// TIA Portal V20 export
Screen "Pop-up_Sealer_1"  395x650
  ScreenItem "Robot Name" at 2,2 size 393x48  Type=HmiIOField
  ScreenItem "Background" at -1,49 size 395x601  Type=HmiRectangle
  ScreenItem "Cancel Mode" at 315,4 size 76x42  Type=HmiButton
  ScreenItem "矩形_4" at 31,68 size 324x517  Type=HmiRectangle
  ScreenItem "Text Filed E- Stop_17" at 39,333 size 148x21  Type=HmiTextBox
  ScreenItem "Text Field In Auto On_9" at 39,98 size 148x21  Type=HmiTextBox
  ScreenItem "Text Field Home Position_17" at 39,121 size 148x21  Type=HmiTextBox
  ScreenItem "Text field Robot Status_5" at 33,69 size 324x26  Type=HmiTextBox
  ScreenItem "Text Field Manual_17" at 39,263 size 148x21  Type=HmiTextBox
  ScreenItem "Text Field System Ready_9" at 39,145 size 148x21  Type=HmiTextBox
  ScreenItem "Text Field Motor On_9" at 39,168 size 148x21  Type=HmiTextBox
  ScreenItem "Text Field In Cycle_9" at 39,192 size 148x21  Type=HmiTextBox
  ScreenItem "Text Field Cycle On_17" at 39,215 size 148x21  Type=HmiTextBox
  ScreenItem "Text Field On Path_17" at 39,239 size 148x21  Type=HmiTextBox
  ScreenItem "Text Field Tryout Mode_17" at 39,286 size 148x21  Type=HmiTextBox
  ScreenItem "Text Field Stop_17" at 39,310 size 148x21  Type=HmiTextBox
  ScreenItem "Text Filed Error_9" at 39,357 size 148x21  Type=HmiTextBox
  ScreenItem "Text Filed Process Fault_9" at 39,380 size 148x21  Type=HmiTextBox
  ScreenItem "Text Field Home Position_18" at 39,404 size 148x21  Type=HmiTextBox
  ScreenItem "Text Filed E- Stop_18" at 39,546 size 148x21  Type=HmiTextBox
  ScreenItem "Text Field Manual_18" at 39,475 size 148x21  Type=HmiTextBox
  ScreenItem "Text Field Cycle On_18" at 39,428 size 148x21  Type=HmiTextBox
  ScreenItem "Text Field On Path_18" at 39,451 size 148x21  Type=HmiTextBox
  ScreenItem "Text Field Tryout Mode_18" at 39,498 size 148x21  Type=HmiTextBox
  ScreenItem "Text Field Stop_18" at 39,522 size 148x21  Type=HmiTextBox
  ScreenItem "Text Filed E- Stop_19" at 200,333 size 148x21  Type=HmiTextBox
  ScreenItem "Text Field In Auto On_10" at 200,98 size 148x21  Type=HmiTextBox
  ScreenItem "Text Field Home Position_19" at 200,121 size 148x21  Type=HmiTextBox
  ScreenItem "Text Field Manual_19" at 200,263 size 148x21  Type=HmiTextBox
  ScreenItem "Text Field System Ready_10" at 200,145 size 148x21  Type=HmiTextBox
  ScreenItem "Text Field Motor On_10" at 200,168 size 148x21  Type=HmiTextBox
  ScreenItem "Text Field In Cycle_10" at 200,192 size 148x21  Type=HmiTextBox
  ScreenItem "Text Field Cycle On_19" at 200,215 size 148x21  Type=HmiTextBox
  ScreenItem "Text Field On Path_19" at 200,239 size 148x21  Type=HmiTextBox
  ScreenItem "Text Field Tryout Mode_19" at 200,286 size 148x21  Type=HmiTextBox
  ScreenItem "Text Field Stop_19" at 200,310 size 148x21  Type=HmiTextBox
  ScreenItem "Text Filed Error_10" at 200,357 size 148x21  Type=HmiTextBox
  ScreenItem "Text Filed Process Fault_10" at 200,380 size 148x21  Type=HmiTextBox
  ScreenItem "Text Field Home Position_20" at 200,404 size 148x21  Type=HmiTextBox
  ScreenItem "Text Filed E- Stop_20" at 200,546 size 148x21  Type=HmiTextBox
  ScreenItem "Text Field Manual_20" at 200,475 size 148x21  Type=HmiTextBox
  ScreenItem "Text Field Cycle On_20" at 200,428 size 148x21  Type=HmiTextBox
  ScreenItem "Text Field On Path_20" at 200,451 size 148x21  Type=HmiTextBox
  ScreenItem "Text Field Tryout Mode_20" at 200,498 size 148x21  Type=HmiTextBox
  ScreenItem "Text Field Stop_20" at 200,522 size 148x21  Type=HmiTextBox
